(* PLC project Vn_fanout_box_to_two_boxes, Beckhoff Automation GmbH TwinCAT PLC Control 3.5.13.21 *)
(* stored: creationDateTime 1970-01-01T00:00:00 *)

PROGRAM Vn_fanout_box_to_two_boxes
  VAR  (* added by the conversion: wires and edge detectors of the diagram *)
    _MAX10000000003_OUT : ANY;
  END_VAR

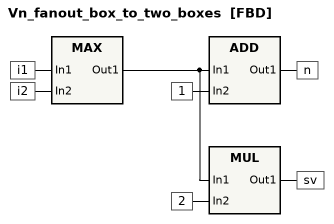
(* FBD diagram, written out as Structured Text *)
_MAX10000000003_OUT := MAX(i1, i2);
n := _MAX10000000003_OUT + 1;
sv := _MAX10000000003_OUT * 2;
END_PROGRAM
